// TIA Portal V21 export
Screen "T13_TplLink"  1024x768, Number=33, Template=Tpl
  ScreenLayer 
    TextField "P_Text" at 0,0 size 100x30  Text="Text"
